// Core S3.8a/S3.8b - the target a manual SET uses (the HMI's operator set
// point): deployment data, never part of a model recipe. SchemaVersion first
// (S3.8b): 0 = never written, 1 = this layout.
TYPE ST_AnalogOutputStationCfg :
STRUCT
    SchemaVersion : UINT;
    ManualTarget  : LREAL;
END_STRUCT
END_TYPE

(* stored: Version 1.1.0.1, ProductVersion 3.1.4024.12
   DUT ST_AnalogOutputStationCfg: Id {6cec4e55-9d26-41f3-8687-c3940c13ecbd} *)
